(* IEC 61131-3 sources: trust-platform/libraries/plant/examples/crusher_lubrication/src, 3 files *)

(* ---- LubricationSequence.st ---- *)
(* Establishes lubrication before the crusher may run: the duty pump runs, then oil flow and
   pressure must be proven within ten seconds; losing either afterwards fails the sequence. The
   sequence commands the pumps through RunPumps, wired to the pump group in Main. *)
USING Plant;

FUNCTION_BLOCK LubricationSequence EXTENDS Plant.FB_Sequence
VAR_INPUT
    PumpRunning : BOOL;
    OilFlow : BOOL;
    Pressure : LREAL;
    MinimumPressure : LREAL := 2.0;
END_VAR
VAR_OUTPUT
    RunPumps : BOOL;
    CrusherPermit : BOOL;
END_VAR
VAR_TEMP
    Proven : BOOL;
END_VAR
    Proven := PumpRunning AND OilFlow AND Pressure >= MinimumPressure;
    IF Execute() THEN
        CASE CurrentStep OF
            0:
                GoTo(Number := 10, Name := 'Establish lubrication');
            10:
                Wait(Text := 'Waiting for a running pump, oil flow and pressure');
                IF Proven THEN
                    GoTo(Number := 20, Name := 'Lubrication ready');
                ELSE
                    StepTimeout(Limit := T#10s, Text := 'Lubrication did not establish within 10 s');
                END_IF;
            20:
                IF NOT Proven THEN
                    Fail(Text := 'Oil flow or pressure lost');
                END_IF;
        END_CASE;
    ELSIF State = E_SequenceState#Stopping THEN
        Wait(Text := 'Stopping the pumps');
        IF NOT PumpRunning THEN
            StopDone();
        END_IF;
    END_IF;
    (* The pumps keep running while the sequence is held; every other state stops them. *)
    RunPumps := State = E_SequenceState#Running OR State = E_SequenceState#Held;
    CrusherPermit := State = E_SequenceState#Running AND CurrentStep = 20;
END_FUNCTION_BLOCK

(* ---- Configuration.st ---- *)
CONFIGURATION Crusher
RESOURCE Cpu ON PLC
    TASK Lubrication (INTERVAL := T#100ms, PRIORITY := 1);
    PROGRAM Application WITH Lubrication : Main;
END_RESOURCE
VAR_CONFIG
    Application.StartButton AT %IX0.0 : BOOL;
    Application.StopButton AT %IX0.1 : BOOL;
    Application.OilLevelOk AT %IX0.2 : BOOL;
    Application.OilFlow AT %IX0.3 : BOOL;
    Application.MainPumpRunning AT %IX0.4 : BOOL;
    Application.StandbyPumpRunning AT %IX0.5 : BOOL;
    Application.MainPumpTrip AT %IX0.6 : BOOL;
    Application.StandbyPumpTrip AT %IX0.7 : BOOL;
    Application.PressureSignal AT %IL1 : LREAL;
    Application.MainPumpRun AT %QX0.0 : BOOL;
    Application.StandbyPumpRun AT %QX0.1 : BOOL;
    Application.CrusherPermit AT %QX0.2 : BOOL;
END_VAR
END_CONFIGURATION

(* ---- Main.st ---- *)
(* Crusher lubrication: two lubrication pumps in a duty/standby group, an oil pressure transmitter,
   an oil level permissive and the lubrication sequence. The pumps run in Auto from the group; an
   operator may take one into Manual from its panel, and the group then uses the other. *)
USING Plant;

PROGRAM Main
VAR
    (* Hardware signals, mapped to I/O in Configuration.st. *)
    StartButton : BOOL;
    StopButton : BOOL;
    OilLevelOk : BOOL;
    OilFlow : BOOL;
    PressureSignal : LREAL;
    MainPumpRunning : BOOL;
    StandbyPumpRunning : BOOL;
    MainPumpTrip : BOOL;
    StandbyPumpTrip : BOOL;
    MainPumpRun : BOOL;
    StandbyPumpRun : BOOL;
    CrusherPermit : BOOL;

    OilPressure : Plant.FB_PressureInput := (Unit := 'bar', RangeHigh := 10.0,
        LowEnabled := TRUE, LowLimit := 1.5, Deadband := 0.1);
    OilLevel : Plant.FB_Permissives;
    MainPump : Plant.FB_Pump;
    StandbyPump : Plant.FB_Pump;
    Pumps : Plant.FB_DutyStandbyGroup := (StartDelay := T#500ms);
    Lubrication : LubricationSequence;
    Alarms : Plant.FB_AlarmManager;
    StartEdge : R_TRIG;
    StopEdge : R_TRIG;
END_VAR
    (* Measurements and conditions first. *)
    OilPressure(Raw := PressureSignal);
    OilLevel(Condition1 := OilLevelOk, Text1 := 'Oil level low');

    (* The push buttons start and stop the sequence; an operator can do the same from its panel. *)
    StartEdge(CLK := StartButton);
    StopEdge(CLK := StopButton);
    IF StartEdge.Q THEN
        Lubrication.Start();
    END_IF;
    IF StopEdge.Q THEN
        Lubrication.Stop();
    END_IF;
    Lubrication(PumpRunning := MainPump.Running OR StandbyPump.Running, OilFlow := OilFlow,
        Pressure := OilPressure.Value);

    (* The group runs one pump while the sequence asks for lubrication; the pumps need oil. *)
    Pumps(Run := Lubrication.RunPumps, Member1 := MainPump, Member2 := StandbyPump);
    MainPump(RunningFeedback := MainPumpRunning, Trip := MainPumpTrip,
        Permissive := OilLevel.Healthy, PermissiveText := OilLevel.Text);
    StandbyPump(RunningFeedback := StandbyPumpRunning, Trip := StandbyPumpTrip,
        Permissive := OilLevel.Healthy, PermissiveText := OilLevel.Text);
    MainPumpRun := MainPump.RunCommand;
    StandbyPumpRun := StandbyPump.RunCommand;
    CrusherPermit := Lubrication.CrusherPermit;

    Alarms(Source1 := MainPump, Source2 := StandbyPump, Source3 := OilPressure, Source4 := Pumps);
END_PROGRAM
